(* PLC project TBEN_L5_PLC11.project, CODESYS CODESYS V3.5 SP21 Patch 1 *)
(* stored: creationDateTime 2026-11-07T15:34:50.7943704, modificationDateTime 2026-11-07T15:09:07.4034196 *)

{attribute 'qualified_only'}
// Quyền truy cập tham số theo IODD (accessRights)
TYPE E_IolAccess :
(
    RO := 0,
    WO := 1,
    RW := 2
) INT;
END_TYPE
